INTERFACE I_LineClamp

METHOD Follow : DINT
VAR_INPUT
    Extend : BOOL;
END_VAR
END_METHOD

METHOD Home
END_METHOD

END_INTERFACE

(* stored: Version 1.1.0.1
   Itf I_LineClamp: Id {CB31703C-BDF0-4A15-AF15-000000000003}
   Method Follow: Id {CB31703C-BDF0-4A15-AF15-000000000001}
   Method Home: Id {CB31703C-BDF0-4A15-AF15-000000000002} *)
